(* Logix 5000 project; controller TFF vendor 1 type 14 code 107 rev 34.11; software revision 34.03; part 34 of 36 *)
(* tags used below, declared in another part *)
   AlarmInhibit_Timer : TIMER;
   Config : Configuration;   // Index Array used in configuration routines
   Index : DINT;   // Index
   NewSystem : DINT;
   SCL : SCALE;   // Scale Instruction
   AlarmAnalog_Storage : AlarmAnalog[6,50];
   AlarmDeviation : AlarmDeviation[20];   // Control Loop Deviation Alarm Array
   AlarmDeviation_Storage : AlarmDeviation[6,20];
   AnalogOutput_Storage : AnalogOutput[6,25];
   AnalogPoint_Storage : AnalogInput[6,50];
   CCPSystem : CCPSystem;   // CCP System Data
   CCPSystem_Storage : CCPSystem_Storage[6];
   ControlLoop : ControlLoop[20];   // Control Loop Array
   ControlLoop_Storage : ControlLoop[6,20];
   DigitalOutput : BOOL[256];   // Digital Output Array these bits are sent to output cards.
   DigitalPoint_Storage : DigitalPoint[6,150];
   Drive : Drive[11];   // Drives Array
   Drive_Storage : Drive[6,11];
   FlowPath : FlowPath[64];   // Flow Path Array
   FlowPath_Storage : FlowPath[6,64];
   LI001 : ALIAS FOR AnalogPoint[44];   // Feed Bag Volume
   LI001Alarm : ALIAS FOR AlarmAnalog[44];   // Feed Bag Volume Alarm
   PCV001_AO : ALIAS FOR AnalogOutput[0];   // Retentate Pressure Control Valve Setpoint
   Phase0 : ALIAS FOR Phase[0];   // Phase 0
   Phase0_Totalizer_Feed : ALIAS FOR PhaseTotalizer[0];   // Phase 0 Total Feed
   PhaseTotalizer_Storage : PhaseTotalizer[6,18];
   PipeAnimation : PipeAnimation;   // HMI Pipe Animation Array
   PSL602 : ALIAS FOR DigitalPoint[0];   // Valves Air Defect
   Rack_Murr_Node1_TF2S : IO_Station;   // Status of Node 1 TF2S
   Rack_Murr_Node1_TF3S : IO_Station;   // Status of Node 1 TF3S
   Rack_Murr_Node4_Instrum_TFF1 : IO_Station;   // Status of Node 4 Instrum TFF1
   Rack_Murr_Node4_Instrum_TFF2 : IO_Station;   // Status of Node 4 Instrum TFF2
   Rack_Murr_Node4_Instrum_TFF3 : IO_Station;   // Status of Node 4 Instrum TFF3
   Rack_Murr_Node4_Instrum_TFF4 : IO_Station;   // Status of Node 4 Instrum TFF4
   Rack_Murr_Node4_Instrum_TFF5 : IO_Station;   // Status of Node 4 Instrum TFF5
   SysControl : SysControl;   // General system status and command
   Tank : TankManagement;   // Tank Management
   ThisSystem : SystemType;
   TI001Alarm : ALIAS FOR AlarmAnalog[13];   // Feed Bag Temperature Alarm
   Valve_Storage : Valve[6,100];
   WI001Alarm : ALIAS FOR AlarmAnalog[15];   // Feed Bag Weight Alarm
   WI101 : ALIAS FOR AnalogPoint[0];   // Filtrate Weight
   WI101Alarm : ALIAS FOR AlarmAnalog[0];   // Filtrate Weight Alarm
   XV001 : ALIAS FOR Valve[0];   // XV001
(* Process, continued *)

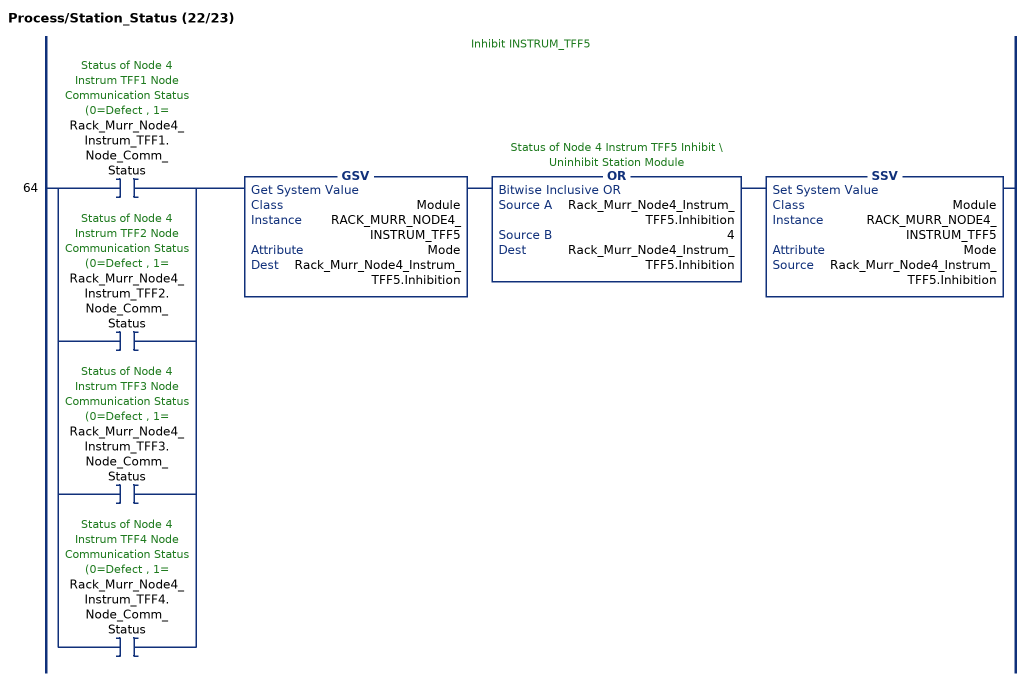
   [picture p431: Process/Station_Status rungs 64-64]
   // Inhibit INSTRUM_TFF5
   64: [XIC(Rack_Murr_Node4_Instrum_TFF1.Node_Comm_Status) ,XIC(Rack_Murr_Node4_Instrum_TFF2.Node_Comm_Status) ,XIC(Rack_Murr_Node4_Instrum_TFF3.Node_Comm_Status) ,XIC(Rack_Murr_Node4_Instrum_TFF4.Node_Comm_Status) ]GSV(Module,RACK_MURR_NODE4_INSTRUM_TFF5,Mode,Rack_Murr_Node4_Instrum_TFF5.Inhibition)OR(Rack_Murr_Node4_Instrum_TFF5.Inhibition,4,Rack_Murr_Node4_Instrum_TFF5.Inhibition)SSV(Module,RACK_MURR_NODE4_INSTRUM_TFF5,Mode,Rack_Murr_Node4_Instrum_TFF5.Inhibition);
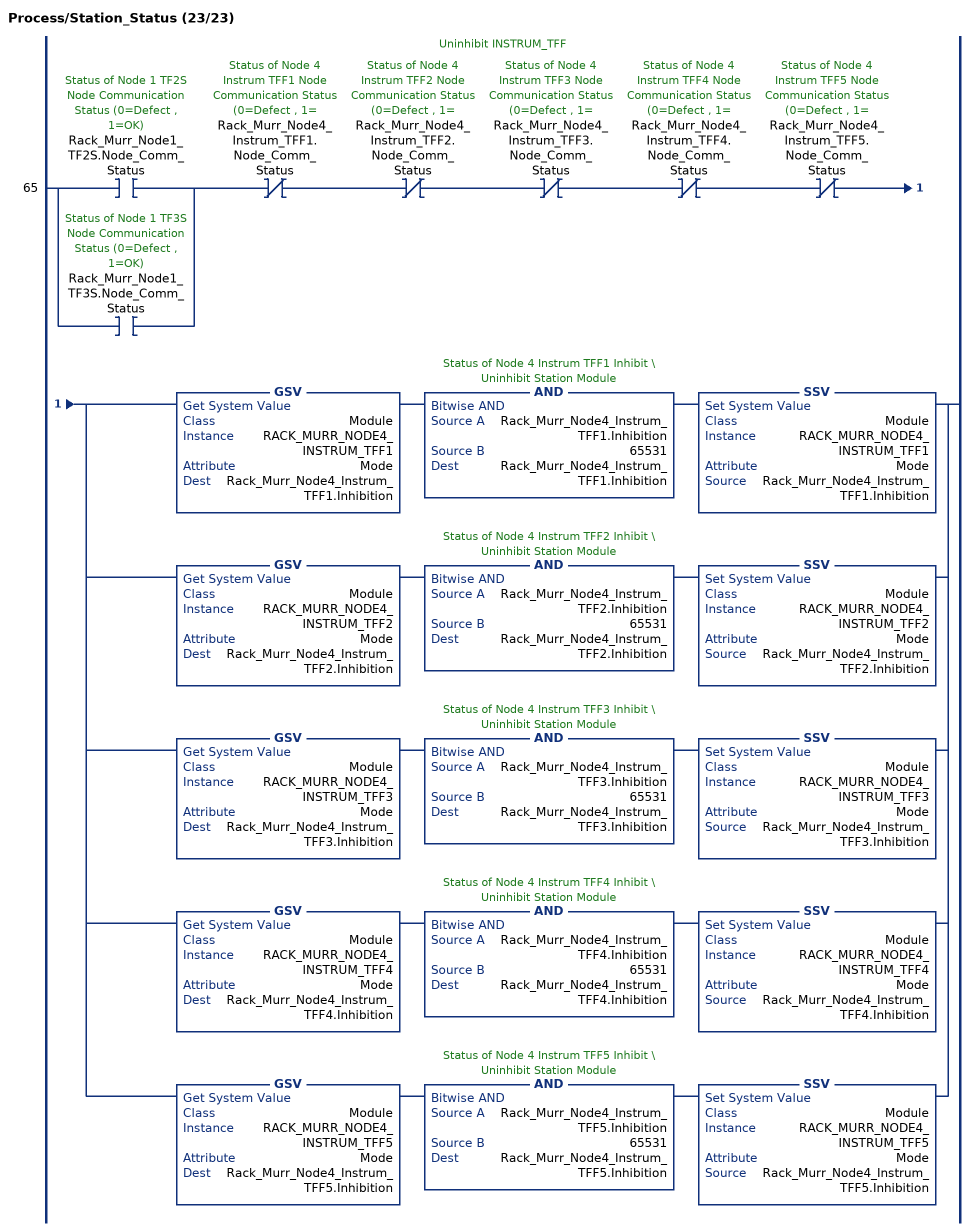
   // Uninhibit INSTRUM_TFF
   65: [XIC(Rack_Murr_Node1_TF2S.Node_Comm_Status) ,XIC(Rack_Murr_Node1_TF3S.Node_Comm_Status) ]XIO(Rack_Murr_Node4_Instrum_TFF1.Node_Comm_Status)XIO(Rack_Murr_Node4_Instrum_TFF2.Node_Comm_Status)XIO(Rack_Murr_Node4_Instrum_TFF3.Node_Comm_Status)XIO(Rack_Murr_Node4_Instrum_TFF4.Node_Comm_Status)XIO(Rack_Murr_Node4_Instrum_TFF5.Node_Comm_Status)[GSV(Module,RACK_MURR_NODE4_INSTRUM_TFF1,Mode,Rack_Murr_Node4_Instrum_TFF1.Inhibition) AND(Rack_Murr_Node4_Instrum_TFF1.Inhibition,65531,Rack_Murr_Node4_Instrum_TFF1.Inhibition) SSV(Module,RACK_MURR_NODE4_INSTRUM_TFF1,Mode,Rack_Murr_Node4_Instrum_TFF1.Inhibition) ,GSV(Module,RACK_MURR_NODE4_INSTRUM_TFF2,Mode,Rack_Murr_Node4_Instrum_TFF2.Inhibition) AND(Rack_Murr_Node4_Instrum_TFF2.Inhibition,65531,Rack_Murr_Node4_Instrum_TFF2.Inhibition) SSV(Module,RACK_MURR_NODE4_INSTRUM_TFF2,Mode,Rack_Murr_Node4_Instrum_TFF2.Inhibition) ,GSV(Module,RACK_MURR_NODE4_INSTRUM_TFF3,Mode,Rack_Murr_Node4_Instrum_TFF3.Inhibition) AND(Rack_Murr_Node4_Instrum_TFF3.Inhibition,65531,Rack_Murr_Node4_Instrum_TFF3.Inhibition) SSV(Module,RACK_MURR_NODE4_INSTRUM_TFF3,Mode,Rack_Murr_Node4_Instrum_TFF3.Inhibition) ,GSV(Module,RACK_MURR_NODE4_INSTRUM_TFF4,Mode,Rack_Murr_Node4_Instrum_TFF4.Inhibition) AND(Rack_Murr_Node4_Instrum_TFF4.Inhibition,65531,Rack_Murr_Node4_Instrum_TFF4.Inhibition) SSV(Module,RACK_MURR_NODE4_INSTRUM_TFF4,Mode,Rack_Murr_Node4_Instrum_TFF4.Inhibition) ,GSV(Module,RACK_MURR_NODE4_INSTRUM_TFF5,Mode,Rack_Murr_Node4_Instrum_TFF5.Inhibition) AND(Rack_Murr_Node4_Instrum_TFF5.Inhibition,65531,Rack_Murr_Node4_Instrum_TFF5.Inhibition) SSV(Module,RACK_MURR_NODE4_INSTRUM_TFF5,Mode,Rack_Murr_Node4_Instrum_TFF5.Inhibition) ];
END_ROUTINE

ROUTINE SystemType   (* ladder *)
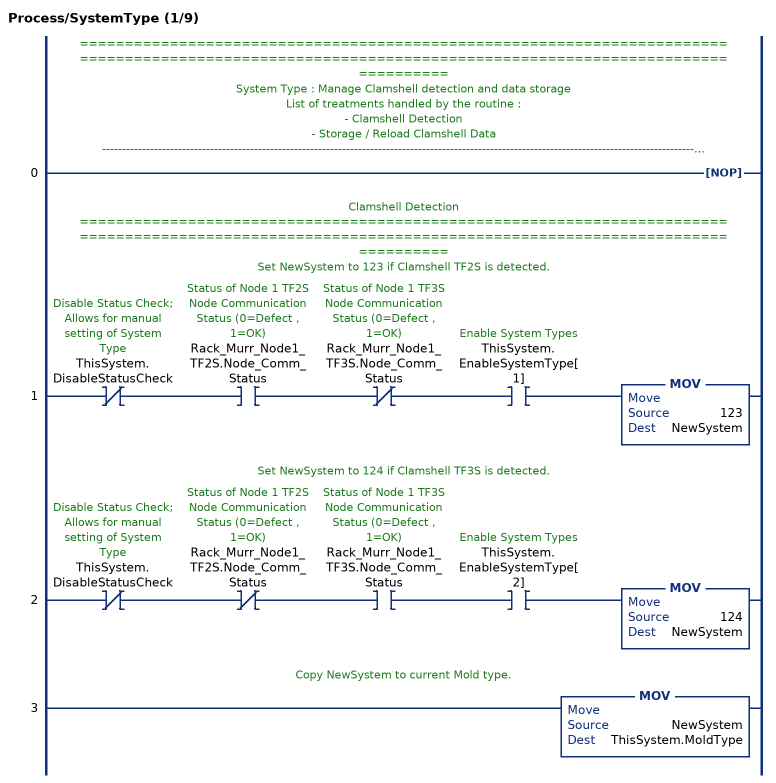
   // ==========================================================================================================================================================
   //                                                               System Type : Manage Clamshell detection and data storage
   //                                                     List of treatments handled by the routine :
   //                                                          - Clamshell Detection
   //                                                          - Storage / Reload Clamshell Data
   //                                                     -----------------------------------------------------------------------------------------------------------------------------------------------------
   //                                                     History
   //                                                          2019-AUG-13 - Actemium - B. Roch - Initial version for Candidate Release 3.00.00.00.a
   // ========================================================================================================================================================
   0: NOP();
   // Clamshell Detection
   // ==========================================================================================================================================================
   // Set NewSystem to 123 if Clamshell TF2S is detected.
   1: XIO(ThisSystem.DisableStatusCheck)XIC(Rack_Murr_Node1_TF2S.Node_Comm_Status)XIO(Rack_Murr_Node1_TF3S.Node_Comm_Status)XIC(ThisSystem.EnableSystemType[1])MOV(123,NewSystem);
   // Set NewSystem to 124 if Clamshell TF3S is detected.
   2: XIO(ThisSystem.DisableStatusCheck)XIO(Rack_Murr_Node1_TF2S.Node_Comm_Status)XIC(Rack_Murr_Node1_TF3S.Node_Comm_Status)XIC(ThisSystem.EnableSystemType[2])MOV(124,NewSystem);
   // Copy NewSystem to current Mold type.
   3: MOV(NewSystem,ThisSystem.MoldType);
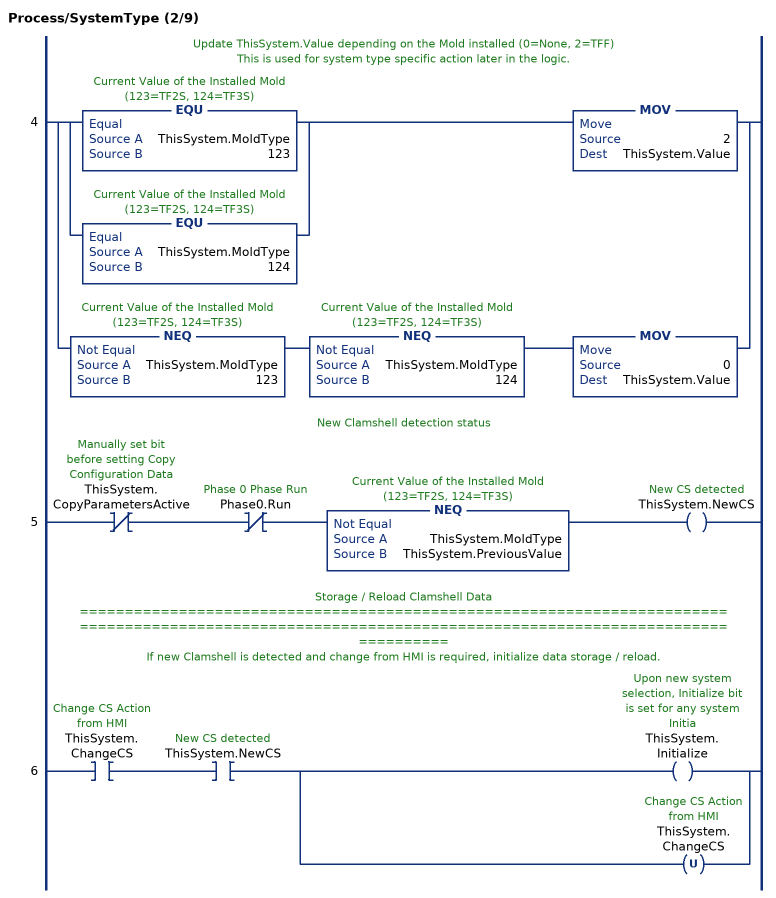
   // Update ThisSystem.Value depending on the Mold installed (0=None, 2=TFF)
   // This is used for system type specific action later in the logic.
   4: [[EQU(ThisSystem.MoldType,123) ,EQU(ThisSystem.MoldType,124) ] MOV(2,ThisSystem.Value) ,NEQ(ThisSystem.MoldType,123) NEQ(ThisSystem.MoldType,124) MOV(0,ThisSystem.Value) ];
   // New Clamshell detection status
   5: XIO(ThisSystem.CopyParametersActive)XIO(Phase0.Run)NEQ(ThisSystem.MoldType,ThisSystem.PreviousValue)OTE(ThisSystem.NewCS);
   // Storage / Reload Clamshell Data
   // ==========================================================================================================================================================
   // If new Clamshell is detected and change from HMI is required, initialize data storage / reload.
   6: XIC(ThisSystem.ChangeCS)XIC(ThisSystem.NewCS)[OTE(ThisSystem.Initialize) ,OTU(ThisSystem.ChangeCS) ];
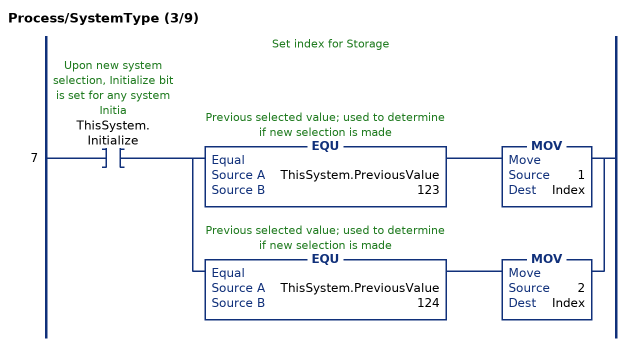
   // Set index for Storage
   7: XIC(ThisSystem.Initialize)[EQU(ThisSystem.PreviousValue,123) MOV(1,Index) ,EQU(ThisSystem.PreviousValue,124) MOV(2,Index) ];
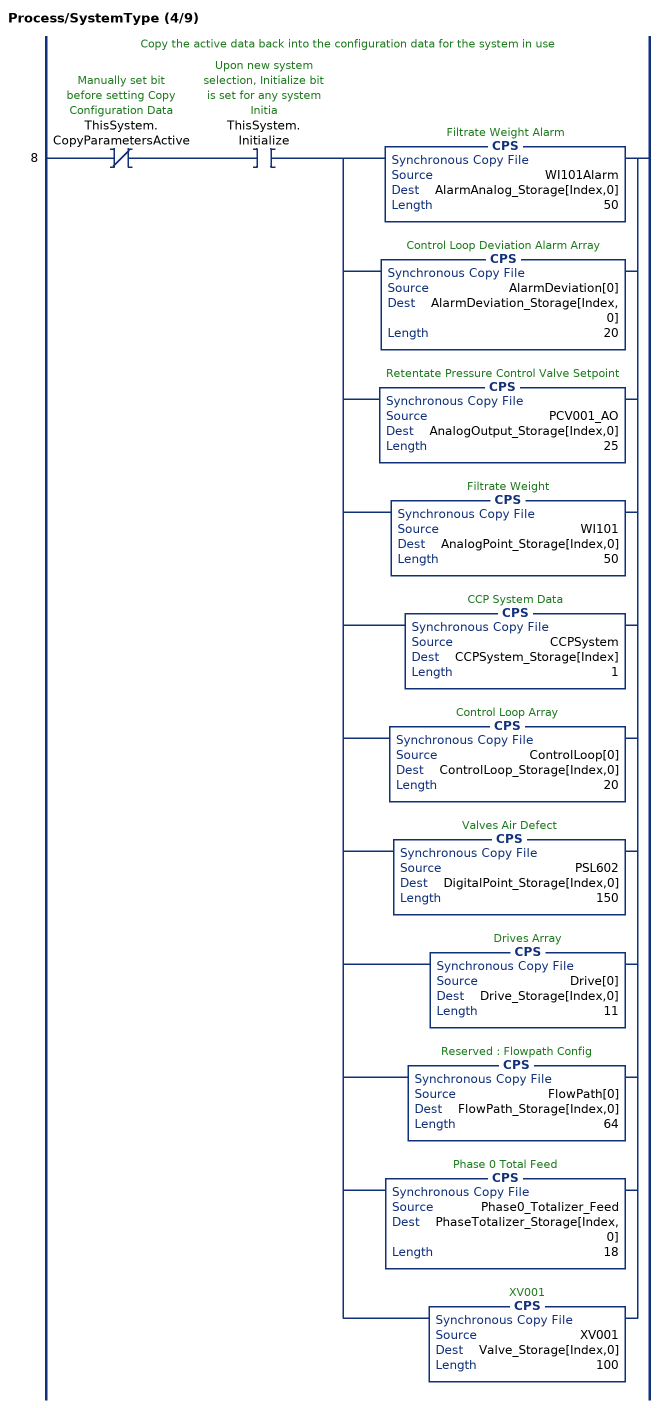
   // Copy the active data back into the configuration data for the system in use
   8: XIO(ThisSystem.CopyParametersActive)XIC(ThisSystem.Initialize)[CPS(WI101Alarm,AlarmAnalog_Storage[Index,0],50) ,CPS(AlarmDeviation[0],AlarmDeviation_Storage[Index,0],20) ,CPS(PCV001_AO,AnalogOutput_Storage[Index,0],25) ,CPS(WI101,AnalogPoint_Storage[Index,0],50) ,CPS(CCPSystem,CCPSystem_Storage[Index],1) ,CPS(ControlLoop[0],ControlLoop_Storage[Index,0],20) ,CPS(PSL602,DigitalPoint_Storage[Index,0],150) ,CPS(Drive[0],Drive_Storage[Index,0],11) ,CPS(FlowPath[0],FlowPath_Storage[Index,0],64) ,CPS(Phase0_Totalizer_Feed,PhaseTotalizer_Storage[Index,0],18) ,CPS(XV001,Valve_Storage[Index,0],100) ];
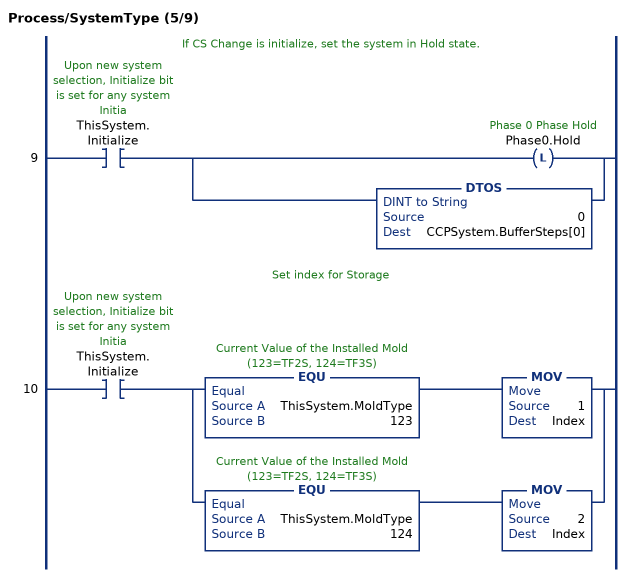
   // If CS Change is initialize, set the system in Hold state.
   9: XIC(ThisSystem.Initialize)[OTL(Phase0.Hold) ,DTOS(0,CCPSystem.BufferSteps[0]) ];
   // Set index for Storage
   10: XIC(ThisSystem.Initialize)[EQU(ThisSystem.MoldType,123) MOV(1,Index) ,EQU(ThisSystem.MoldType,124) MOV(2,Index) ];
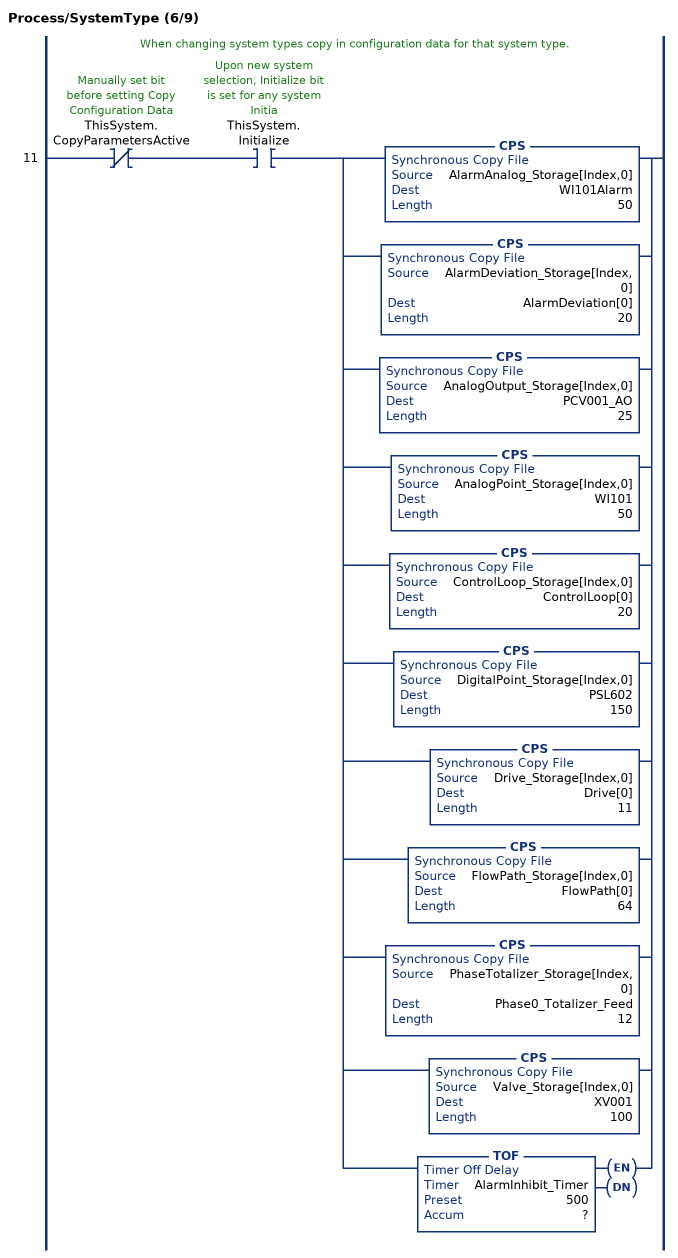
   // When changing system types copy in configuration data for that system type.
   11: XIO(ThisSystem.CopyParametersActive)XIC(ThisSystem.Initialize)[CPS(AlarmAnalog_Storage[Index,0],WI101Alarm,50) ,CPS(AlarmDeviation_Storage[Index,0],AlarmDeviation[0],20) ,CPS(AnalogOutput_Storage[Index,0],PCV001_AO,25) ,CPS(AnalogPoint_Storage[Index,0],WI101,50) ,CPS(ControlLoop_Storage[Index,0],ControlLoop[0],20) ,CPS(DigitalPoint_Storage[Index,0],PSL602,150) ,CPS(Drive_Storage[Index,0],Drive[0],11) ,CPS(FlowPath_Storage[Index,0],FlowPath[0],64) ,CPS(PhaseTotalizer_Storage[Index,0],Phase0_Totalizer_Feed,12) ,CPS(Valve_Storage[Index,0],XV001,100) ,TOF(AlarmInhibit_Timer,?,?) ];
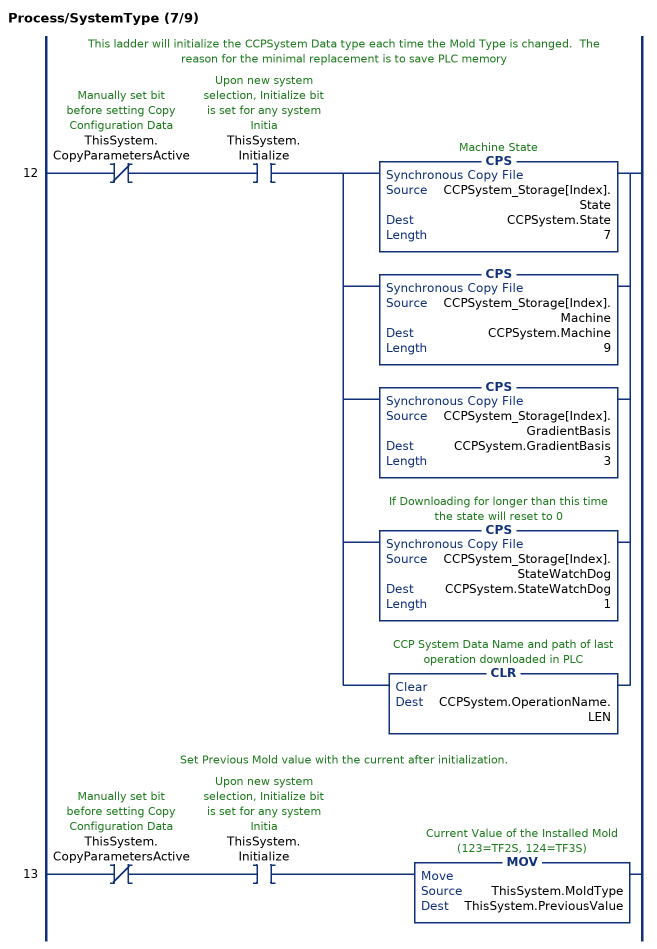
   // This ladder will initialize the CCPSystem Data type each time the Mold Type is changed.  The reason for the minimal replacement is to save PLC memory
   12: XIO(ThisSystem.CopyParametersActive)XIC(ThisSystem.Initialize)[CPS(CCPSystem_Storage[Index].State,CCPSystem.State,7) ,CPS(CCPSystem_Storage[Index].Machine,CCPSystem.Machine,9) ,CPS(CCPSystem_Storage[Index].GradientBasis,CCPSystem.GradientBasis,3) ,CPS(CCPSystem_Storage[Index].StateWatchDog,CCPSystem.StateWatchDog,1) ,CLR(CCPSystem.OperationName.LEN) ];
   // Set Previous Mold value with the current after initialization.
   13: XIO(ThisSystem.CopyParametersActive)XIC(ThisSystem.Initialize)MOV(ThisSystem.MoldType,ThisSystem.PreviousValue);
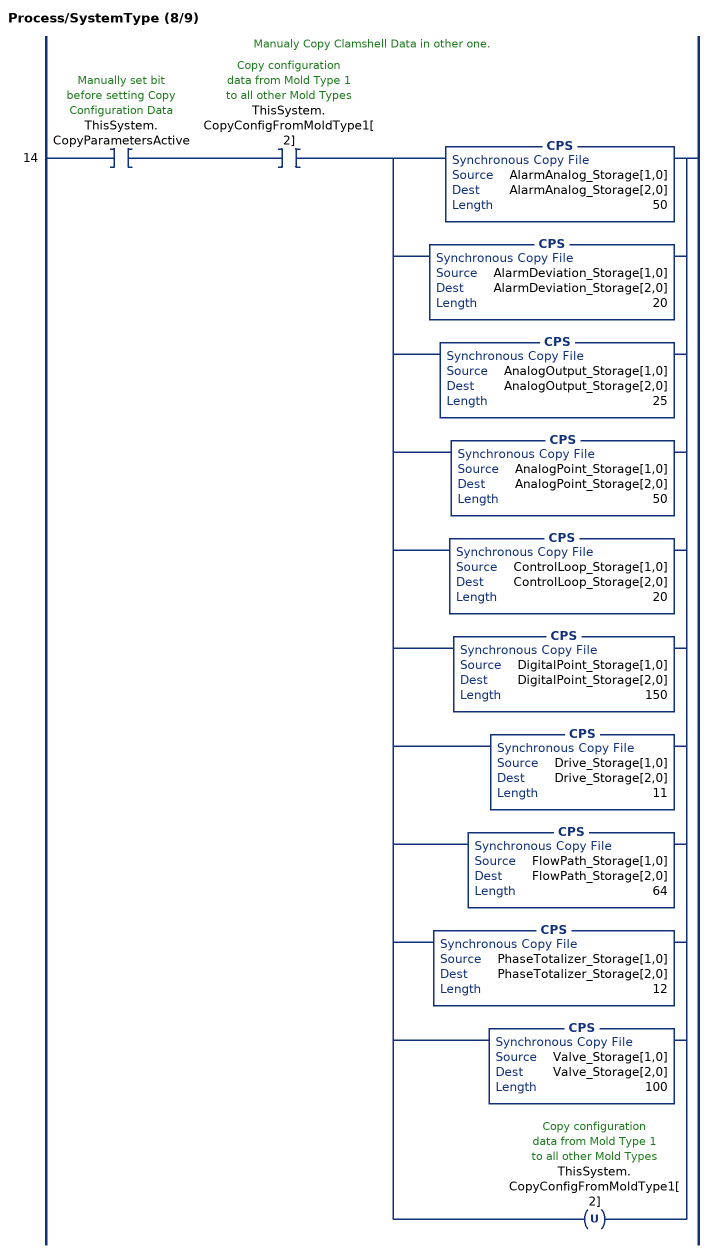
   // Manualy Copy Clamshell Data in other one.
   14: XIC(ThisSystem.CopyParametersActive)XIC(ThisSystem.CopyConfigFromMoldType1[2])[CPS(AlarmAnalog_Storage[1,0],AlarmAnalog_Storage[2,0],50) ,CPS(AlarmDeviation_Storage[1,0],AlarmDeviation_Storage[2,0],20) ,CPS(AnalogOutput_Storage[1,0],AnalogOutput_Storage[2,0],25) ,CPS(AnalogPoint_Storage[1,0],AnalogPoint_Storage[2,0],50) ,CPS(ControlLoop_Storage[1,0],ControlLoop_Storage[2,0],20) ,CPS(DigitalPoint_Storage[1,0],DigitalPoint_Storage[2,0],150) ,CPS(Drive_Storage[1,0],Drive_Storage[2,0],11) ,CPS(FlowPath_Storage[1,0],FlowPath_Storage[2,0],64) ,CPS(PhaseTotalizer_Storage[1,0],PhaseTotalizer_Storage[2,0],12) ,CPS(Valve_Storage[1,0],Valve_Storage[2,0],100) ,OTU(ThisSystem.CopyConfigFromMoldType1[2]) ];
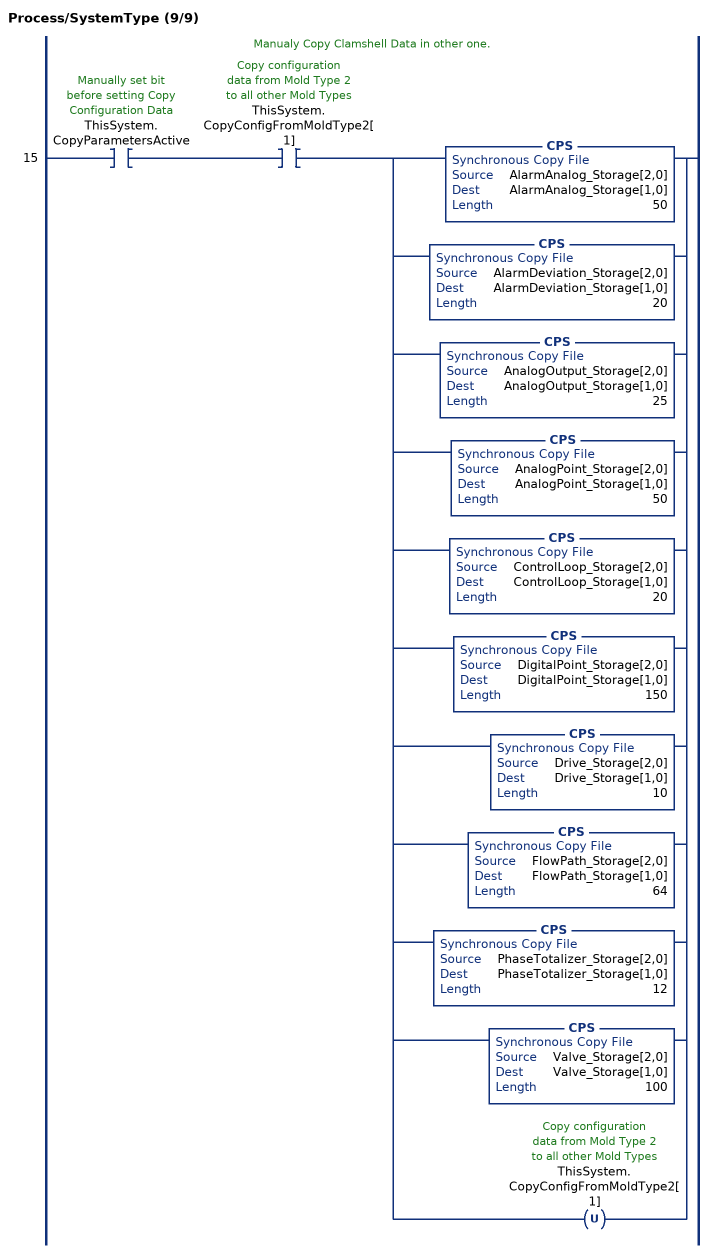
   // Manualy Copy Clamshell Data in other one.
   15: XIC(ThisSystem.CopyParametersActive)XIC(ThisSystem.CopyConfigFromMoldType2[1])[CPS(AlarmAnalog_Storage[2,0],AlarmAnalog_Storage[1,0],50) ,CPS(AlarmDeviation_Storage[2,0],AlarmDeviation_Storage[1,0],20) ,CPS(AnalogOutput_Storage[2,0],AnalogOutput_Storage[1,0],25) ,CPS(AnalogPoint_Storage[2,0],AnalogPoint_Storage[1,0],50) ,CPS(ControlLoop_Storage[2,0],ControlLoop_Storage[1,0],20) ,CPS(DigitalPoint_Storage[2,0],DigitalPoint_Storage[1,0],150) ,CPS(Drive_Storage[2,0],Drive_Storage[1,0],10) ,CPS(FlowPath_Storage[2,0],FlowPath_Storage[1,0],64) ,CPS(PhaseTotalizer_Storage[2,0],PhaseTotalizer_Storage[1,0],12) ,CPS(Valve_Storage[2,0],Valve_Storage[1,0],100) ,OTU(ThisSystem.CopyConfigFromMoldType2[1]) ];
END_ROUTINE

ROUTINE TankManagement   (* ladder *)
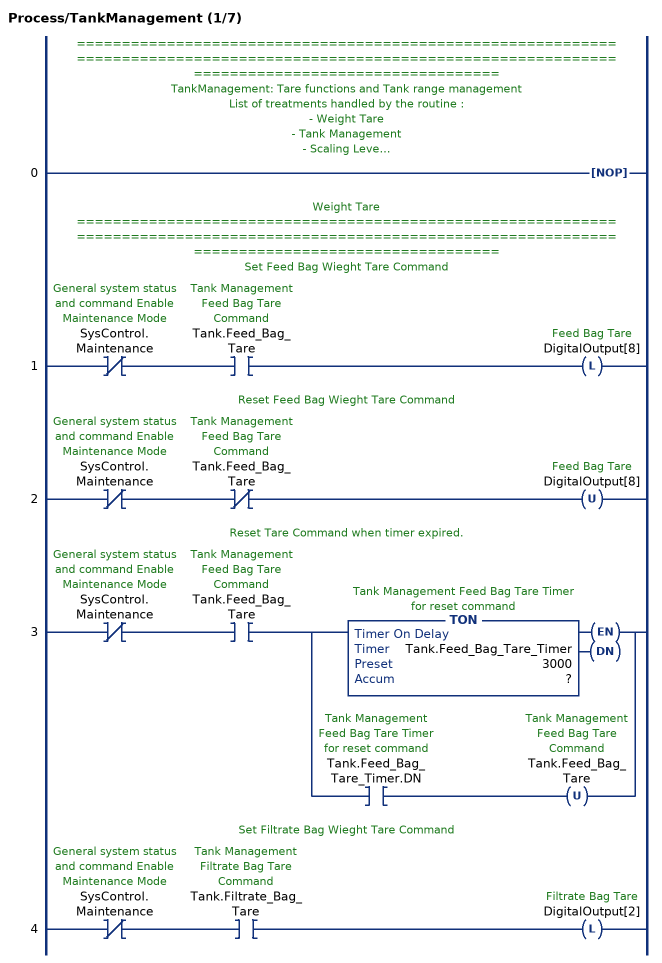
   // ==========================================================================================================================================================
   //                                                                                                                                 TankManagement: Tare functions and Tank range management
   //                                                     List of treatments handled by the routine :
   //                                                          - Weight Tare
   //                                                          - Tank Management
   //                                                          - Scaling Level
   //                                                          - Tank Status
   //                                                     -----------------------------------------------------------------------------------------------------------------------------------------------------
   //                                                     History
   //                                                          2019-AUG-13 - Actemium - B. Roch - Initial version for Candidate Release 3.00.00.00.a
   // ==========================================================================================================================================================
   0: NOP();
   // Weight Tare
   // ==========================================================================================================================================================
   // Set Feed Bag Wieght Tare Command
   1: XIO(SysControl.Maintenance)XIC(Tank.Feed_Bag_Tare)OTL(DigitalOutput[8]);
   // Reset Feed Bag Wieght Tare Command
   2: XIO(SysControl.Maintenance)XIO(Tank.Feed_Bag_Tare)OTU(DigitalOutput[8]);
   // Reset Tare Command when timer expired.
   3: XIO(SysControl.Maintenance)XIC(Tank.Feed_Bag_Tare)[TON(Tank.Feed_Bag_Tare_Timer,?,?) ,XIC(Tank.Feed_Bag_Tare_Timer.DN) OTU(Tank.Feed_Bag_Tare) ];
   // Set Filtrate Bag Wieght Tare Command
   4: XIO(SysControl.Maintenance)XIC(Tank.Filtrate_Bag_Tare)OTL(DigitalOutput[2]);
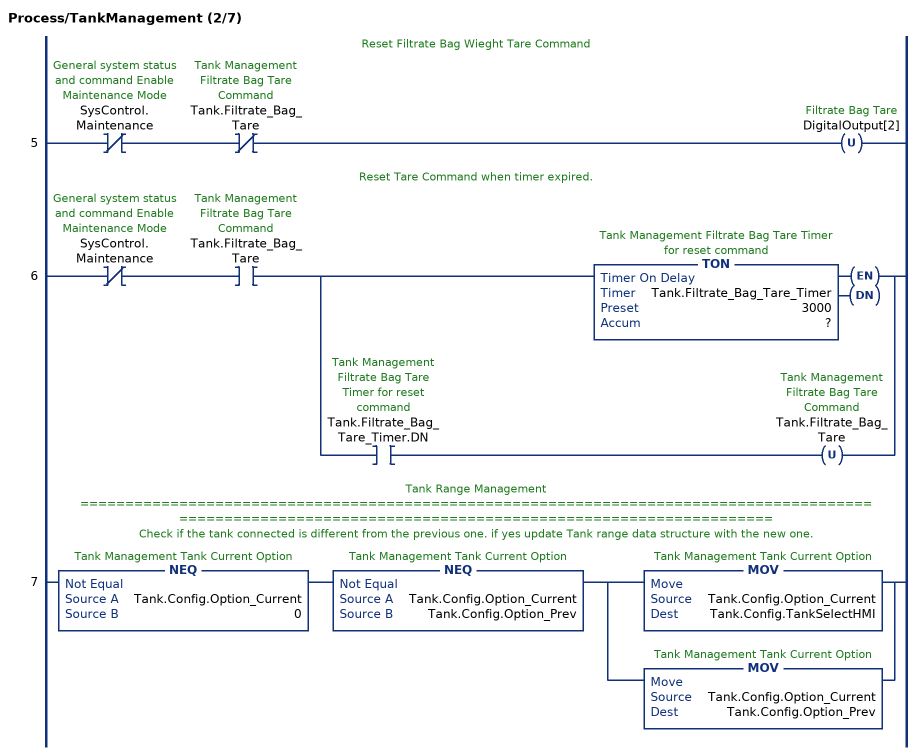
   // Reset Filtrate Bag Wieght Tare Command
   5: XIO(SysControl.Maintenance)XIO(Tank.Filtrate_Bag_Tare)OTU(DigitalOutput[2]);
   // Reset Tare Command when timer expired.
   6: XIO(SysControl.Maintenance)XIC(Tank.Filtrate_Bag_Tare)[TON(Tank.Filtrate_Bag_Tare_Timer,?,?) ,XIC(Tank.Filtrate_Bag_Tare_Timer.DN) OTU(Tank.Filtrate_Bag_Tare) ];
   // Tank Range Management
   // ==========================================================================================================================================================
   // Check if the tank connected is different from the previous one. if yes update Tank range data structure with the new one.
   7: NEQ(Tank.Config.Option_Current,0)NEQ(Tank.Config.Option_Current,Tank.Config.Option_Prev)[MOV(Tank.Config.Option_Current,Tank.Config.TankSelectHMI) ,MOV(Tank.Config.Option_Current,Tank.Config.Option_Prev) ];
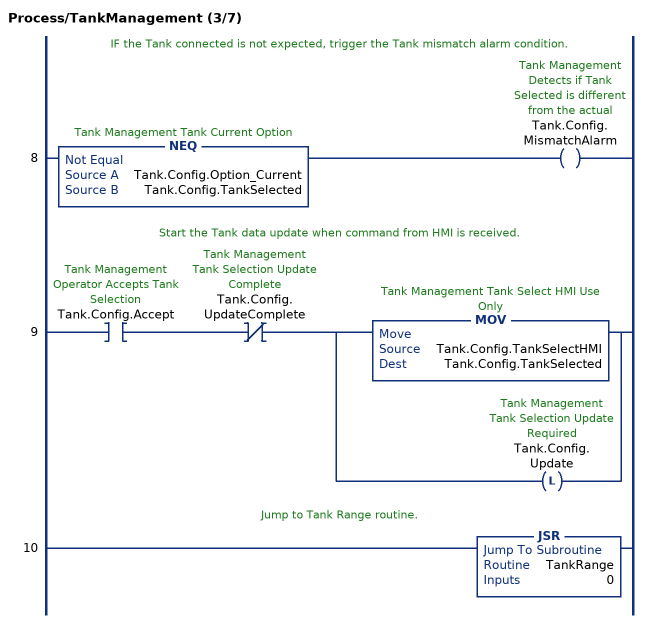
   // IF the Tank connected is not expected, trigger the Tank mismatch alarm condition.
   8: NEQ(Tank.Config.Option_Current,Tank.Config.TankSelected)OTE(Tank.Config.MismatchAlarm);
   // Start the Tank data update when command from HMI is received.
   9: XIC(Tank.Config.Accept)XIO(Tank.Config.UpdateComplete)[MOV(Tank.Config.TankSelectHMI,Tank.Config.TankSelected) ,OTL(Tank.Config.Update) ];
   // Jump to Tank Range routine.
   10: JSR(TankRange,0);
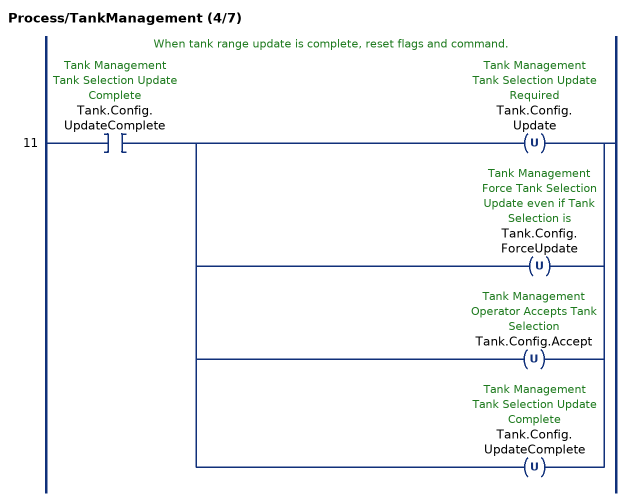
   // When tank range update is complete, reset flags and command.
   11: XIC(Tank.Config.UpdateComplete)[OTU(Tank.Config.Update) ,OTU(Tank.Config.ForceUpdate) ,OTU(Tank.Config.Accept) ,OTU(Tank.Config.UpdateComplete) ];
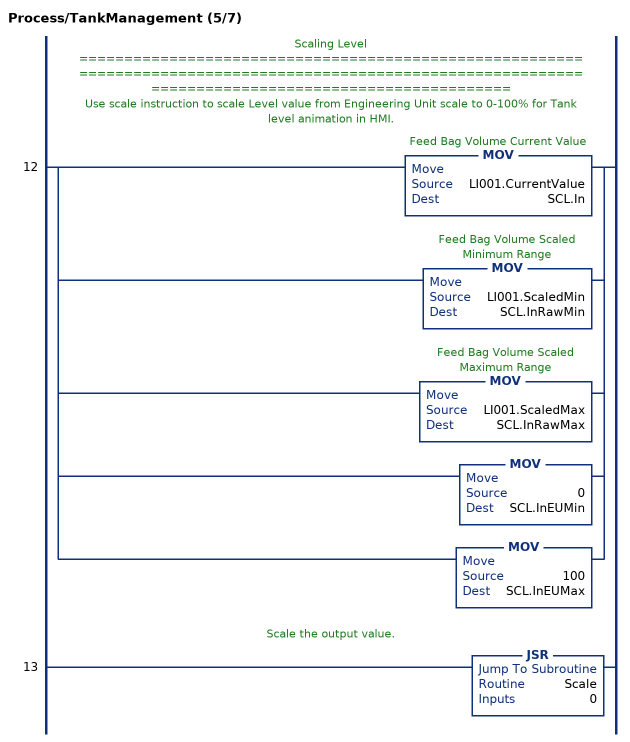
   // Scaling Level
   // ========================================================================================================================================================
   // Use scale instruction to scale Level value from Engineering Unit scale to 0-100% for Tank level animation in HMI.
   12: [MOV(LI001.CurrentValue,SCL.In) ,MOV(LI001.ScaledMin,SCL.InRawMin) ,MOV(LI001.ScaledMax,SCL.InRawMax) ,MOV(0,SCL.InEUMin) ,MOV(100,SCL.InEUMax) ];
   // Scale the output value.
   13: JSR(Scale,0);
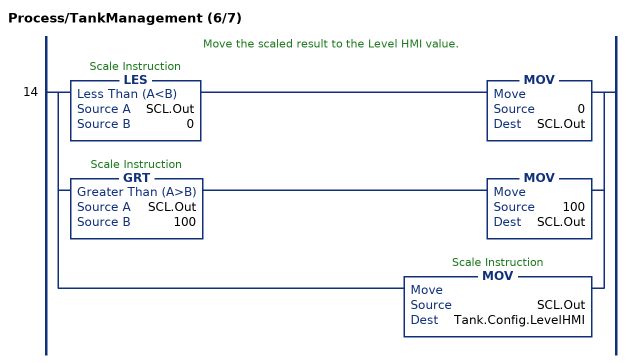
   // Move the scaled result to the Level HMI value.
   14: [LES(SCL.Out,0) MOV(0,SCL.Out) ,GRT(SCL.Out,100) MOV(100,SCL.Out) ,MOV(SCL.Out,Tank.Config.LevelHMI) ];
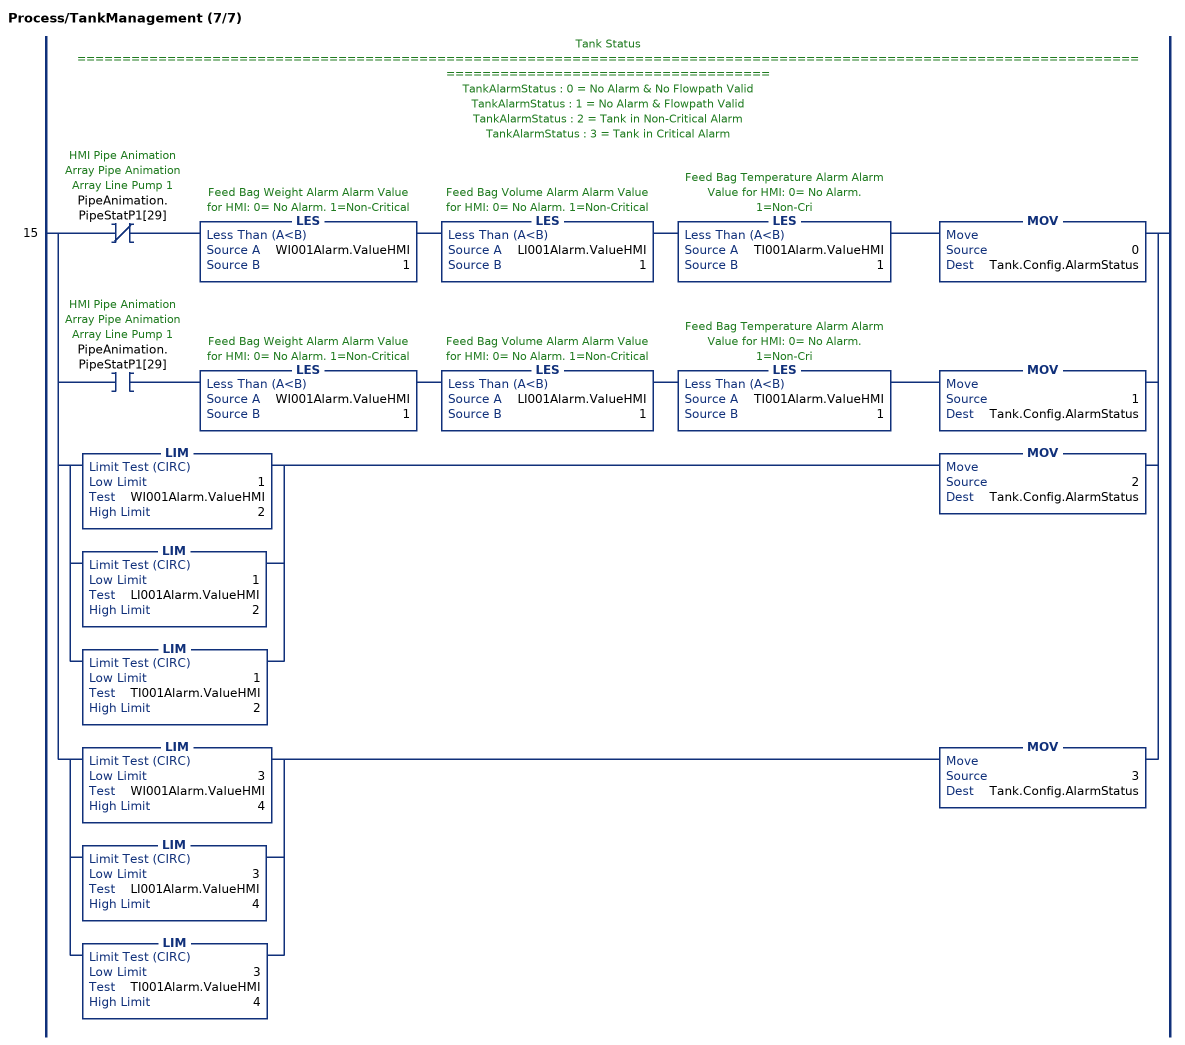
   // Tank Status
   // ==========================================================================================================================================================
   // TankAlarmStatus : 0 = No Alarm & No Flowpath Valid
   // TankAlarmStatus : 1 = No Alarm & Flowpath Valid
   // TankAlarmStatus : 2 = Tank in Non-Critical Alarm
   // TankAlarmStatus : 3 = Tank in Critical Alarm
   15: [XIO(PipeAnimation.PipeStatP1[29]) LES(WI001Alarm.ValueHMI,1) LES(LI001Alarm.ValueHMI,1) LES(TI001Alarm.ValueHMI,1) MOV(0,Tank.Config.AlarmStatus) ,XIC(PipeAnimation.PipeStatP1[29]) LES(WI001Alarm.ValueHMI,1) LES(LI001Alarm.ValueHMI,1) LES(TI001Alarm.ValueHMI,1) MOV(1,Tank.Config.AlarmStatus) ,[LIM(1,WI001Alarm.ValueHMI,2) ,LIM(1,LI001Alarm.ValueHMI,2) ,LIM(1,TI001Alarm.ValueHMI,2) ] MOV(2,Tank.Config.AlarmStatus) ,[LIM(3,WI001Alarm.ValueHMI,4) ,LIM(3,LI001Alarm.ValueHMI,4) ,LIM(3,TI001Alarm.ValueHMI,4) ] MOV(3,Tank.Config.AlarmStatus) ];
END_ROUTINE
